TYPE "ST_FraktalHal"
VERSION : 0.1
   STRUCT
      "PressDemo" {ExternalAccessible := 'False'; ExternalVisible := 'False'; ExternalWritable := 'False'} : "ST_PressDemoUnitHal";
   END_STRUCT;
END_TYPE
